FUNCTION_BLOCK FB_RParamInit
VAR_INPUT
	bExecute	:	BOOL	:=	FALSE;
END_VAR
VAR_OUTPUT
	bBusy		:	BOOL	:=	FALSE;
	bErr		:	BOOL	:=	FALSE;
END_VAR
VAR_IN_OUT
	inst_NcToPlc_NCI	:	NCTOPLC_NCICHANNEL_REF;
END_VAR
VAR
	BusyIdx		:	DINT	:=	0;	
	nState		:	DINT	:=	0;
	fb_WriteRParams	:	ItpWriteRParams;
END_VAR

CASE nState OF
	
0:
	IF bExecute THEN
		bBusy	:=	TRUE;
		bErr	:=	FALSE;
		nState	:=	1;
		BusyIdx	:=	0;
	END_IF

1:
	fb_WriteRParams(
		bExecute	:=	TRUE,
		nChnId		:=	inst_NcToPlc_NCI.ChnId,
		pAddr		:=	ADR(UserVar.R_InitVal),
		nIndex		:=	TO_DINT(UserVar.R_Params[BusyIdx]),
		nCount		:=	1);
	nState	:=	2;


2:
	IF fb_WriteRParams.bBusy THEN
		fb_WriteRParams(
			bExecute	:=	FALSE,
			nChnId		:=	inst_NcToPlc_NCI.ChnId,
			pAddr		:=	ADR(UserVar.R_InitVal),
			nIndex		:=	TO_DINT(UserVar.R_Params[BusyIdx]),
			nCount		:=	1);
		nState	:=	3;
	END_IF
	

3:	
	fb_WriteRParams(	bExecute	:=	FALSE);
	IF NOT fb_WriteRParams.bBusy THEN
		IF fb_WriteRParams.bErr THEN
			bErr	:=	TRUE;
			bBusy	:=	FALSE;
			nState	:=	0;
		ELSE
			BusyIdx	:=	BusyIdx	+	1;
			IF BusyIdx 	>=	(SIZEOF(UserVar.R_Params) / 2) THEN
				bBusy	:=	FALSE;
				nState	:=	0;
			ELSE
				nState	:=	1;
			END_IF
		END_IF
	END_IF

END_CASE

END_FUNCTION_BLOCK

(* stored: Version 1.1.0.1, ProductVersion 3.1.4024.15
   POU FB_RParamInit: Id {1fba08f7-68e7-45dd-8820-debf83ddb4b9}, SpecialFunc None *)
